Fanuc KAREL source: compact_preamble.KL

PROGRAM KX00023
%NOLOCKGROUP
VAR
I:INTEGER;J:INTEGER;B:BOOLEAN
F : FILE
S : STRING[80]
P : XYZWPR
PE : XYZWPREXT
BEGIN
PE.X=1.0
P=PE
END KX00023
